% RSLogix 500 project LadderLogicforProject_Rslogix500file.RSS, saved by version 8.40.00.08 %
PROJECT "UNTITLED"    % processor: MicroLogix 1400 %

PROGRAM FILES
  LAD 2   7 rungs

DATA FILES
  O0 OUTPUT  6 elements
  I1 INPUT  8 elements
  S2 STATUS  66 elements
  B3 BINARY  1 elements
  T4 TIMER  1 elements
  C5 COUNTER  1 elements
  R6 CONTROL  1 elements
  N7 INTEGER  1 elements
  F8 FLOAT  1 elements

LADDER 2
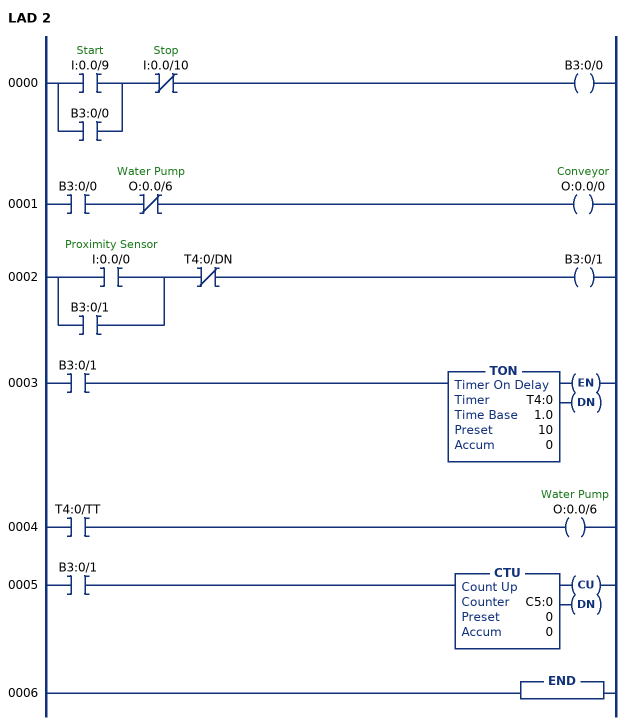
% Rung: 0 %
SOR BST XIC I:0.0/9 NXB XIC B3:0/0 BND XIO I:0.0/10 OTE B3:0/0 EOR
%   I:0.0/9  "Start" %
%   I:0.0/10  "Stop" %
% Rung: 1 %
SOR XIC B3:0/0 XIO O:0.0/6 OTE O:0.0/0 EOR
%   O:0.0/6  "Water Pump" %
%   O:0.0/0  "Conveyor" %
% Rung: 2 %
SOR BST XIC I:0.0/0 NXB XIC B3:0/1 BND XIO T4:0/DN OTE B3:0/1 EOR
%   I:0.0/0  "Proximity Sensor" %
% Rung: 3 %
SOR XIC B3:0/1 TON T4:0 1.0 10 0 EOR
% Rung: 4 %
SOR XIC T4:0/TT OTE O:0.0/6 EOR
%   O:0.0/6  "Water Pump" %
% Rung: 5 %
SOR XIC B3:0/1 CTU C5:0 0 0 EOR
% Rung: 6 %
SOR END EOR

OTHER DOCUMENTED ADDRESSES
  I:0.0/1  "Stop"
  I:0.0/2  "Proximity Sensor"
  O:0.0/1  "Water Pump"

DATA TABLE (non-zero values as saved)
DATA T4
% .PRE .ACC %
% T4:0 % 10 0
